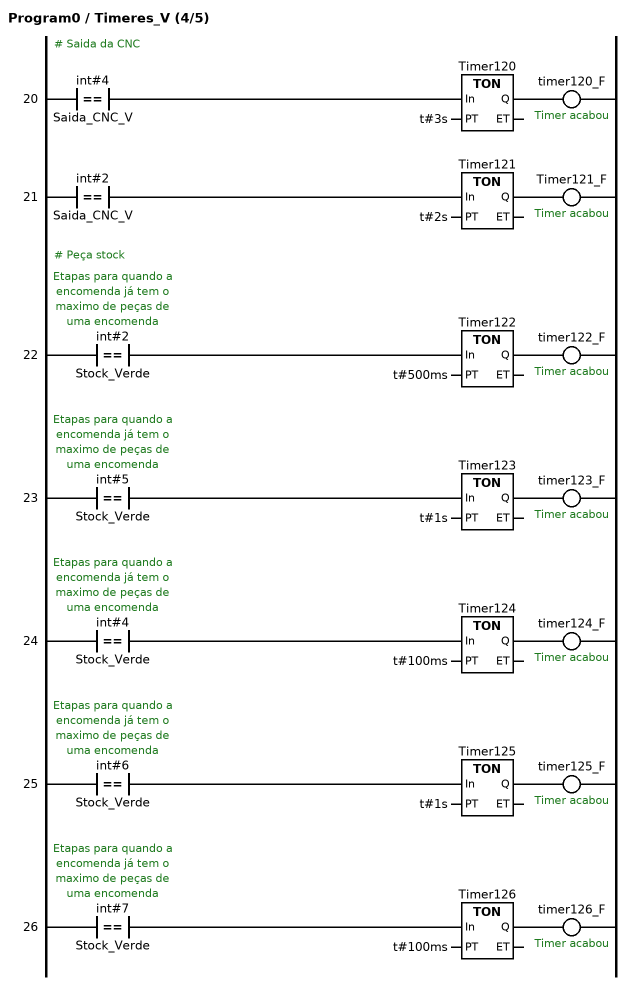
(* [picture p24: Program0 / Timeres_V, rungs 20-26] *)
(* Rung 20: # Saida da CNC *)
Timer120(In := int#4 = Saida_CNC_V, PT := t#3s);
timer120_F := Timer120.Q;
(* Rung 21 *)
Timer121(In := int#2 = Saida_CNC_V, PT := t#2s);
Timer121_F := Timer121.Q;
(* Rung 22: # Peça stock *)
Timer122(In := int#2 = Stock_Verde, PT := t#500ms);
timer122_F := Timer122.Q;
(* Rung 23 *)
Timer123(In := int#5 = Stock_Verde, PT := t#1s);
timer123_F := Timer123.Q;
(* Rung 24 *)
Timer124(In := int#4 = Stock_Verde, PT := t#100ms);
timer124_F := Timer124.Q;
(* Rung 25 *)
Timer125(In := int#6 = Stock_Verde, PT := t#1s);
timer125_F := Timer125.Q;
(* Rung 26 *)
Timer126(In := int#7 = Stock_Verde, PT := t#100ms);
timer126_F := Timer126.Q;

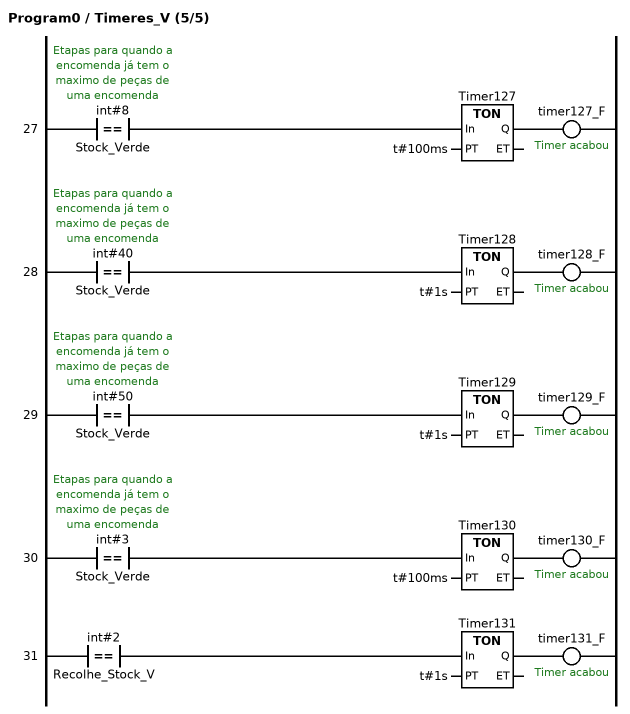
(* Rung 27 *)
Timer127(In := int#8 = Stock_Verde, PT := t#100ms);
timer127_F := Timer127.Q;
(* Rung 28 *)
Timer128(In := int#40 = Stock_Verde, PT := t#1s);
timer128_F := Timer128.Q;
(* Rung 29 *)
Timer129(In := int#50 = Stock_Verde, PT := t#1s);
timer129_F := Timer129.Q;
(* Rung 30 *)
Timer130(In := int#3 = Stock_Verde, PT := t#100ms);
timer130_F := Timer130.Q;
(* Rung 31 *)
Timer131(In := int#2 = Recolhe_Stock_V, PT := t#1s);
timer131_F := Timer131.Q;

(* Section Timeres_C: ladder, written here as Structured Text *)

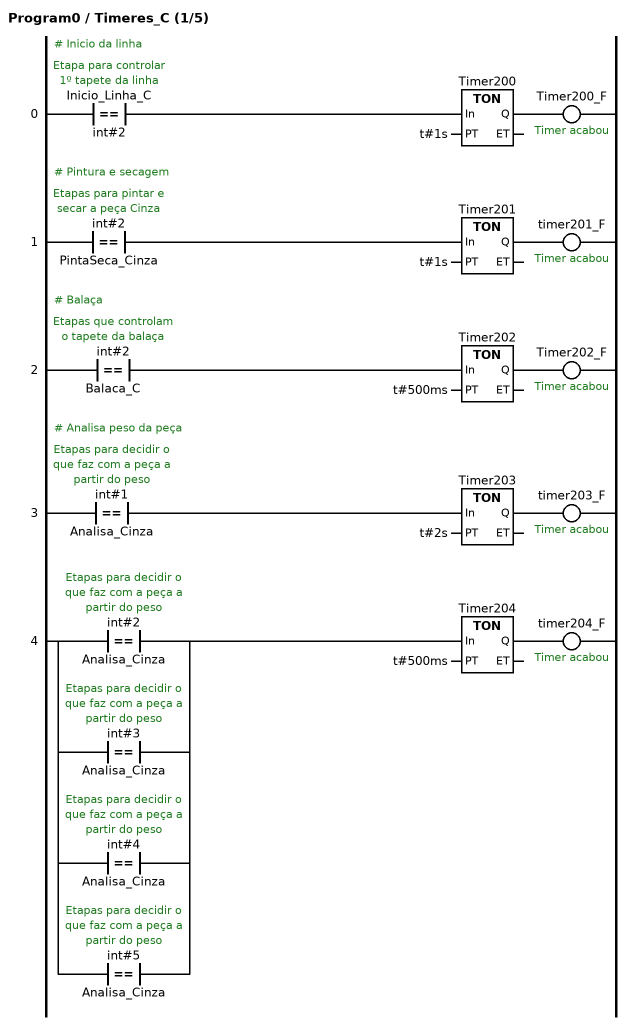
(* Rung 0: # Inicio da linha *)
Timer200(In := Inicio_Linha_C = int#2, PT := t#1s);
Timer200_F := Timer200.Q;
(* Rung 1: # Pintura e secagem *)
Timer201(In := int#2 = PintaSeca_Cinza, PT := t#1s);
timer201_F := Timer201.Q;
(* Rung 2: # Balaça *)
Timer202(In := int#2 = Balaca_C, PT := t#500ms);
Timer202_F := Timer202.Q;
(* Rung 3: # Analisa peso da peça *)
Timer203(In := int#1 = Analisa_Cinza, PT := t#2s);
timer203_F := Timer203.Q;
(* Rung 4 *)
Timer204(In := (int#2 = Analisa_Cinza) OR (int#3 = Analisa_Cinza) OR (int#4 = Analisa_Cinza) OR (int#5 = Analisa_Cinza), PT := t#500ms);
timer204_F := Timer204.Q;

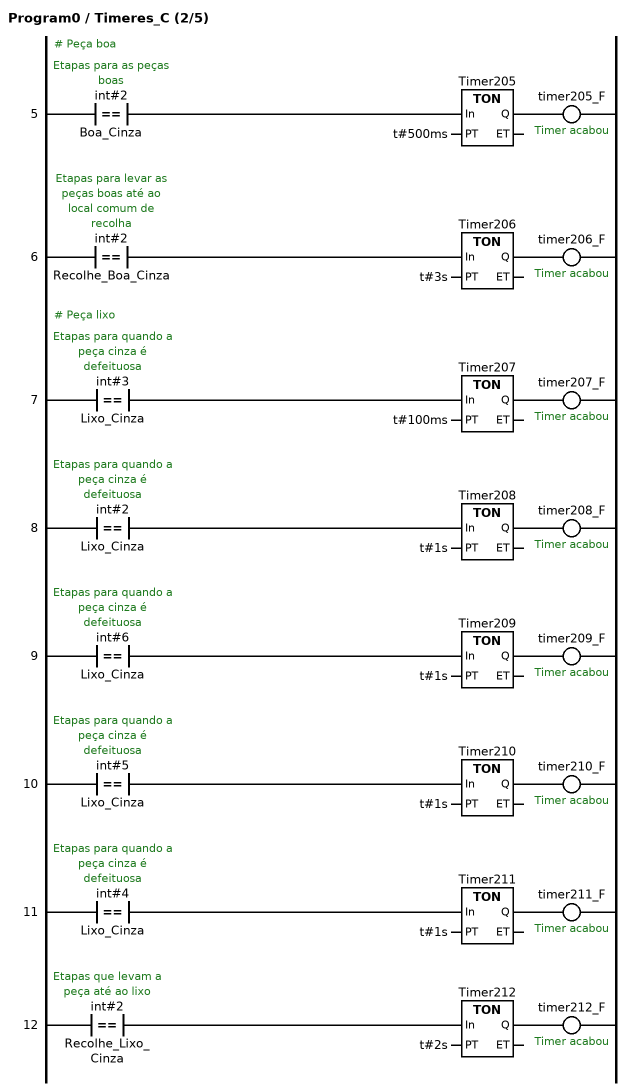
(* Rung 5: # Peça boa *)
Timer205(In := int#2 = Boa_Cinza, PT := t#500ms);
timer205_F := Timer205.Q;
(* Rung 6 *)
Timer206(In := int#2 = Recolhe_Boa_Cinza, PT := t#3s);
timer206_F := Timer206.Q;
(* Rung 7: # Peça lixo *)
Timer207(In := int#3 = Lixo_Cinza, PT := t#100ms);
timer207_F := Timer207.Q;
(* Rung 8 *)
Timer208(In := int#2 = Lixo_Cinza, PT := t#1s);
timer208_F := Timer208.Q;
(* Rung 9 *)
Timer209(In := int#6 = Lixo_Cinza, PT := t#1s);
timer209_F := Timer209.Q;
(* Rung 10 *)
Timer210(In := int#5 = Lixo_Cinza, PT := t#1s);
timer210_F := Timer210.Q;
(* Rung 11 *)
Timer211(In := int#4 = Lixo_Cinza, PT := t#1s);
timer211_F := Timer211.Q;
(* Rung 12 *)
Timer212(In := int#2 = Recolhe_Lixo_Cinza, PT := t#2s);
timer212_F := Timer212.Q;

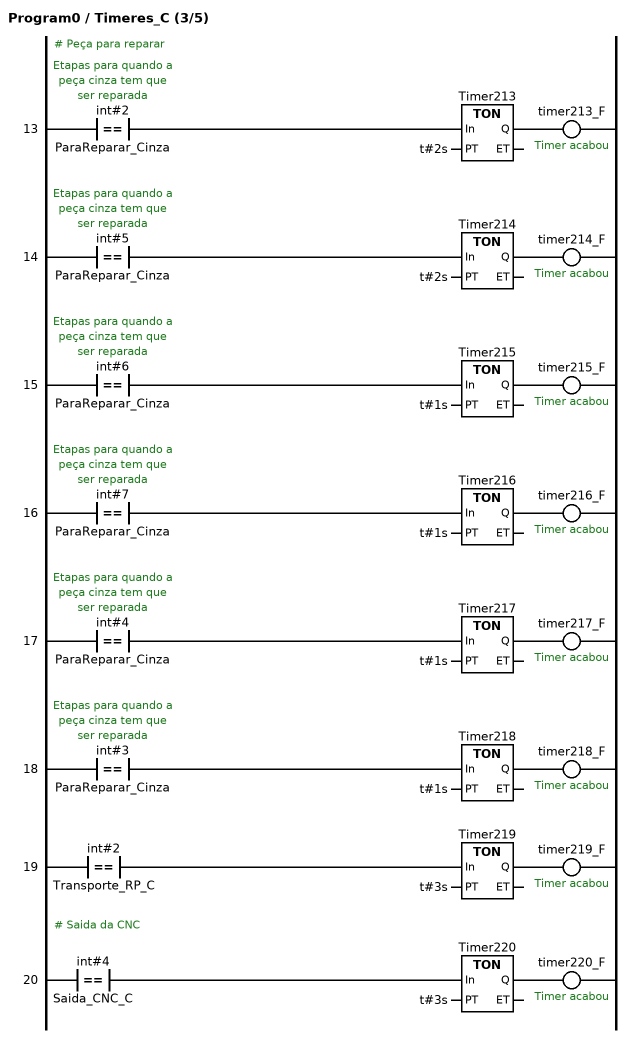
(* Rung 13: # Peça para reparar *)
Timer213(In := int#2 = ParaReparar_Cinza, PT := t#2s);
timer213_F := Timer213.Q;
(* Rung 14 *)
Timer214(In := int#5 = ParaReparar_Cinza, PT := t#2s);
timer214_F := Timer214.Q;
(* Rung 15 *)
Timer215(In := int#6 = ParaReparar_Cinza, PT := t#1s);
timer215_F := Timer215.Q;
(* Rung 16 *)
Timer216(In := int#7 = ParaReparar_Cinza, PT := t#1s);
timer216_F := Timer216.Q;
(* Rung 17 *)
Timer217(In := int#4 = ParaReparar_Cinza, PT := t#1s);
timer217_F := Timer217.Q;
(* Rung 18 *)
Timer218(In := int#3 = ParaReparar_Cinza, PT := t#1s);
timer218_F := Timer218.Q;
(* Rung 19 *)
Timer219(In := int#2 = Transporte_RP_C, PT := t#3s);
timer219_F := Timer219.Q;
(* Rung 20: # Saida da CNC *)
Timer220(In := int#4 = Saida_CNC_C, PT := t#3s);
timer220_F := Timer220.Q;

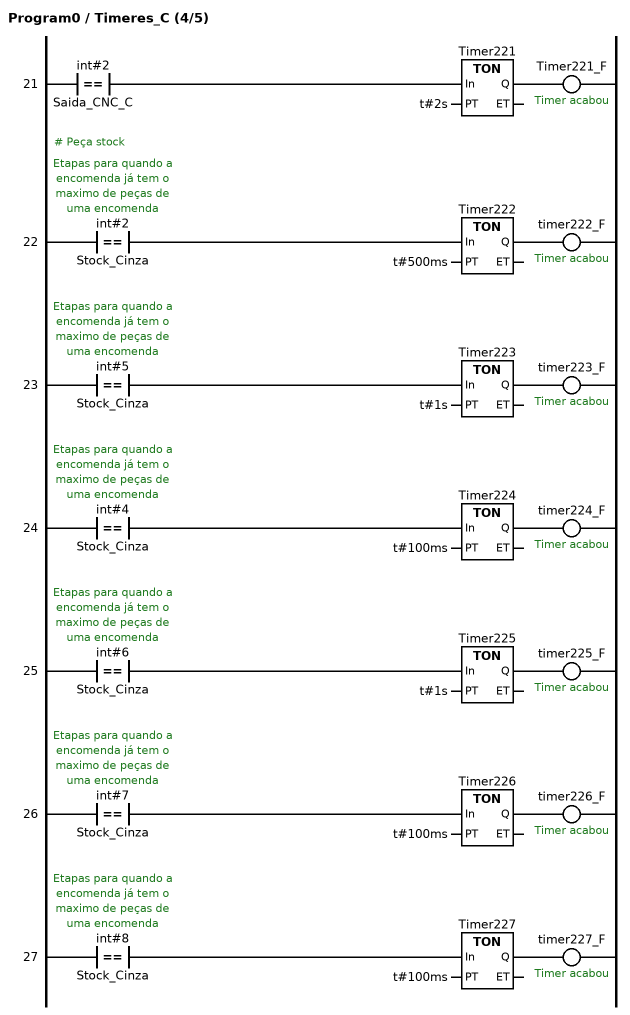
(* Rung 21 *)
Timer221(In := int#2 = Saida_CNC_C, PT := t#2s);
Timer221_F := Timer221.Q;
(* Rung 22: # Peça stock *)
Timer222(In := int#2 = Stock_Cinza, PT := t#500ms);
timer222_F := Timer222.Q;
(* Rung 23 *)
Timer223(In := int#5 = Stock_Cinza, PT := t#1s);
timer223_F := Timer223.Q;
(* Rung 24 *)
Timer224(In := int#4 = Stock_Cinza, PT := t#100ms);
timer224_F := Timer224.Q;
(* Rung 25 *)
Timer225(In := int#6 = Stock_Cinza, PT := t#1s);
timer225_F := Timer225.Q;
(* Rung 26 *)
Timer226(In := int#7 = Stock_Cinza, PT := t#100ms);
timer226_F := Timer226.Q;
(* Rung 27 *)
Timer227(In := int#8 = Stock_Cinza, PT := t#100ms);
timer227_F := Timer227.Q;

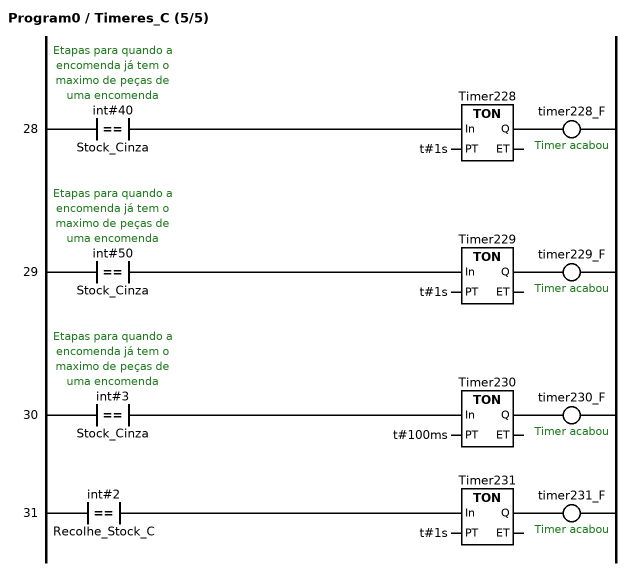
(* Rung 28 *)
Timer228(In := int#40 = Stock_Cinza, PT := t#1s);
timer228_F := Timer228.Q;
(* Rung 29 *)
Timer229(In := int#50 = Stock_Cinza, PT := t#1s);
timer229_F := Timer229.Q;
(* Rung 30 *)
Timer230(In := int#3 = Stock_Cinza, PT := t#100ms);
timer230_F := Timer230.Q;
(* Rung 31 *)
Timer231(In := int#2 = Recolhe_Stock_C, PT := t#1s);
timer231_F := Timer231.Q;

(* Section Emitter_Removers: ladder, written here as Structured Text *)

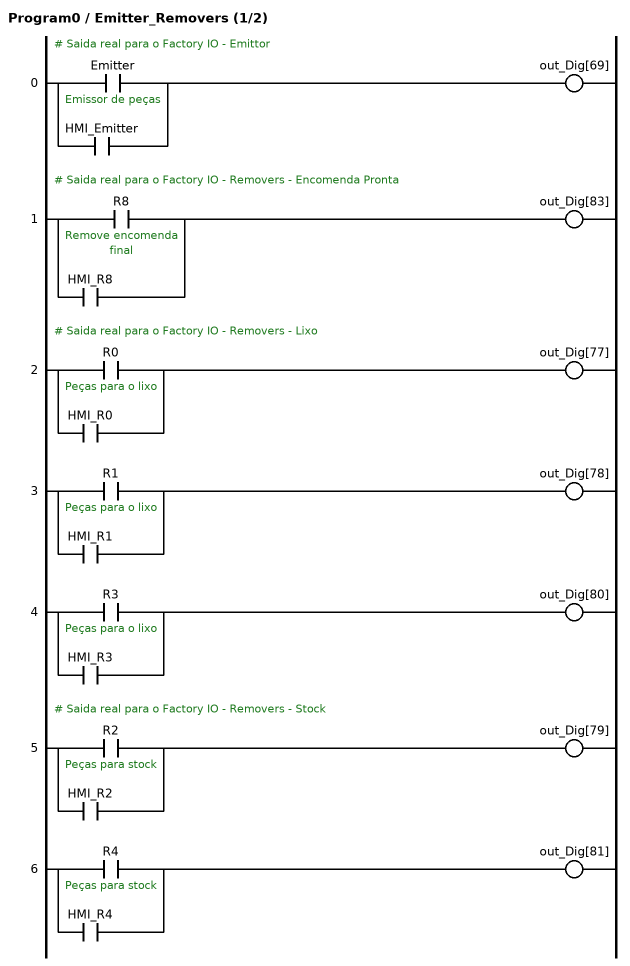
(* Rung 0: # Saida real para o Factory IO - Emittor *)
out_Dig[69] := Emitter OR HMI_Emitter;
(* Rung 1: # Saida real para o Factory IO - Removers - Encomenda Pronta *)
out_Dig[83] := R8 OR HMI_R8;
(* Rung 2: # Saida real para o Factory IO - Removers - Lixo *)
out_Dig[77] := R0 OR HMI_R0;
(* Rung 3 *)
out_Dig[78] := R1 OR HMI_R1;
(* Rung 4 *)
out_Dig[80] := R3 OR HMI_R3;
(* Rung 5: # Saida real para o Factory IO - Removers - Stock *)
out_Dig[79] := R2 OR HMI_R2;
(* Rung 6 *)
out_Dig[81] := R4 OR HMI_R4;

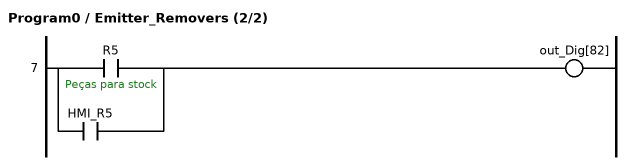
(* Rung 7 *)
out_Dig[82] := R5 OR HMI_R5;

(* Section Semaforos_Alarme: ladder, written here as Structured Text *)

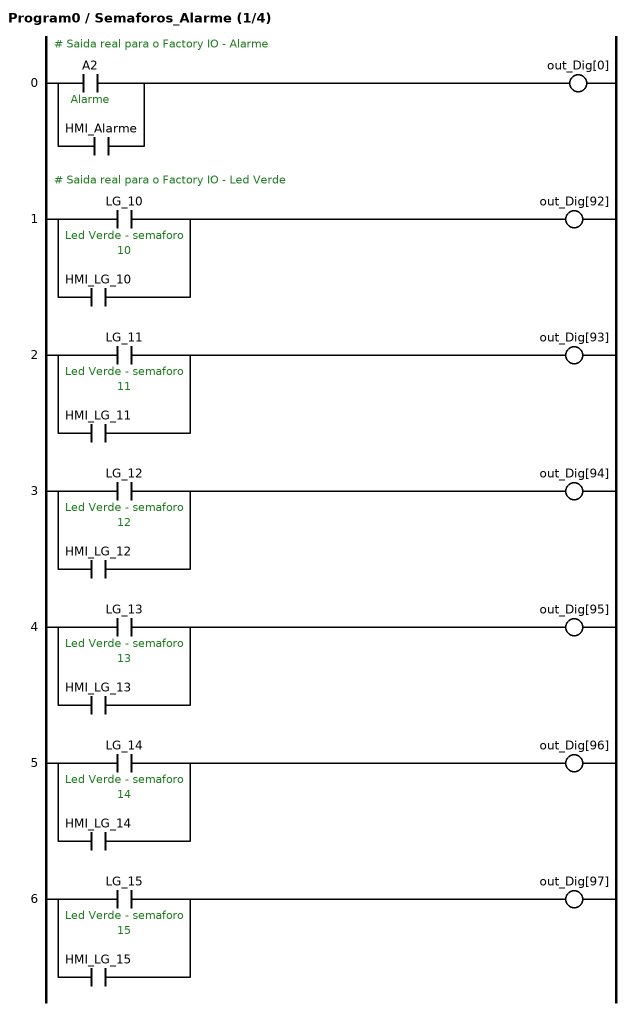
(* Rung 0: # Saida real para o Factory IO - Alarme *)
out_Dig[0] := A2 OR HMI_Alarme;
(* Rung 1: # Saida real para o Factory IO - Led Verde *)
out_Dig[92] := LG_10 OR HMI_LG_10;
(* Rung 2 *)
out_Dig[93] := LG_11 OR HMI_LG_11;
(* Rung 3 *)
out_Dig[94] := LG_12 OR HMI_LG_12;
(* Rung 4 *)
out_Dig[95] := LG_13 OR HMI_LG_13;
(* Rung 5 *)
out_Dig[96] := LG_14 OR HMI_LG_14;
(* Rung 6 *)
out_Dig[97] := LG_15 OR HMI_LG_15;

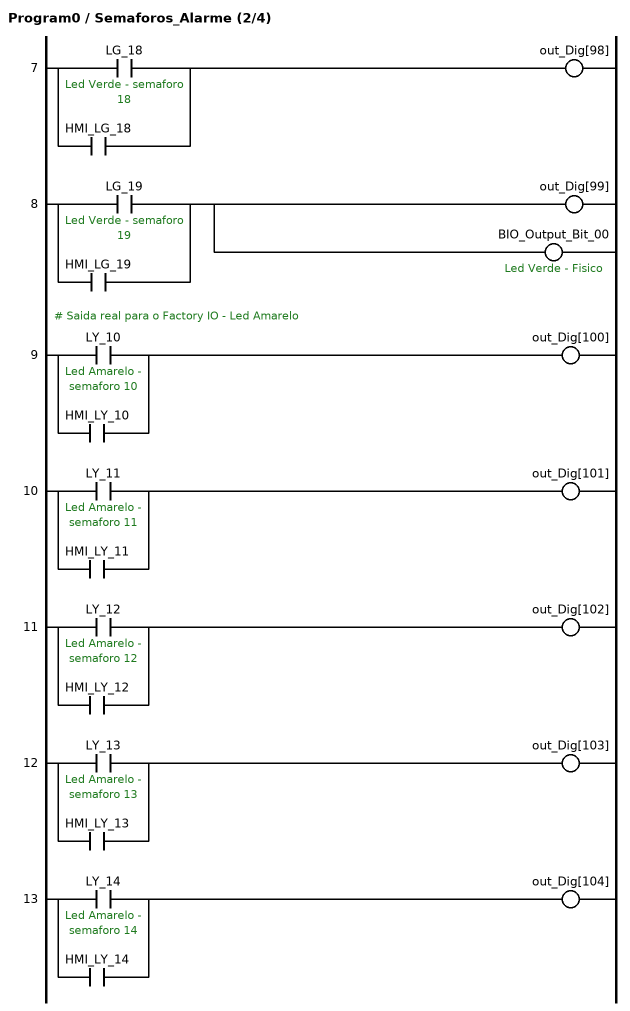
(* Rung 7 *)
out_Dig[98] := LG_18 OR HMI_LG_18;
(* Rung 8 *)
out_Dig[99] := LG_19 OR HMI_LG_19;
BIO_Output_Bit_00 := LG_19 OR HMI_LG_19;
(* Rung 9: # Saida real para o Factory IO - Led Amarelo *)
out_Dig[100] := LY_10 OR HMI_LY_10;
(* Rung 10 *)
out_Dig[101] := LY_11 OR HMI_LY_11;
(* Rung 11 *)
out_Dig[102] := LY_12 OR HMI_LY_12;
(* Rung 12 *)
out_Dig[103] := LY_13 OR HMI_LY_13;
(* Rung 13 *)
out_Dig[104] := LY_14 OR HMI_LY_14;

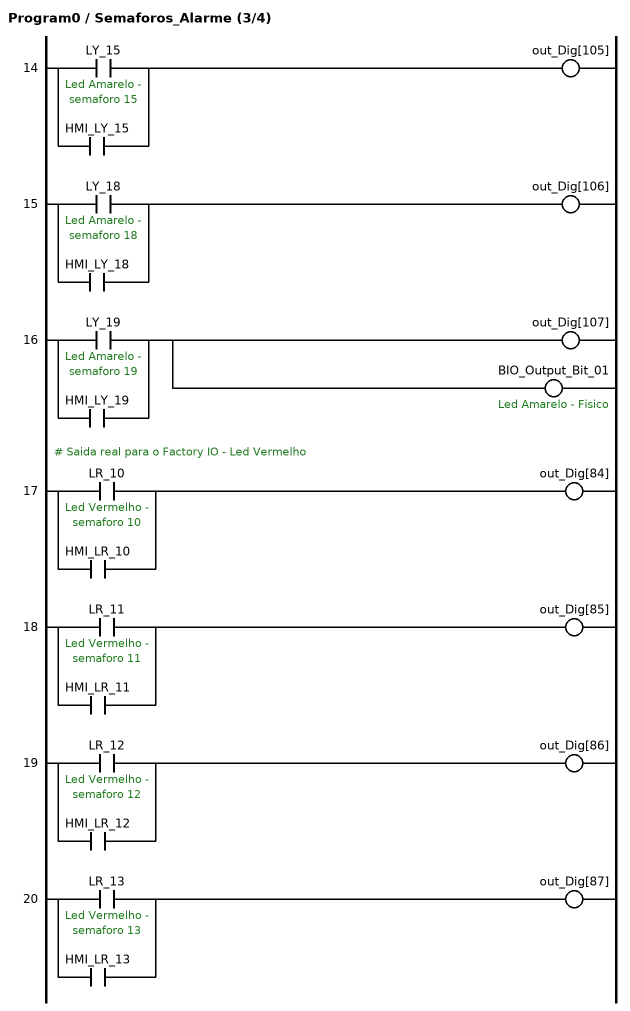
(* Rung 14 *)
out_Dig[105] := LY_15 OR HMI_LY_15;
(* Rung 15 *)
out_Dig[106] := LY_18 OR HMI_LY_18;
(* Rung 16 *)
out_Dig[107] := LY_19 OR HMI_LY_19;
BIO_Output_Bit_01 := LY_19 OR HMI_LY_19;
(* Rung 17: # Saida real para o Factory IO - Led Vermelho *)
out_Dig[84] := LR_10 OR HMI_LR_10;
(* Rung 18 *)
out_Dig[85] := LR_11 OR HMI_LR_11;
(* Rung 19 *)
out_Dig[86] := LR_12 OR HMI_LR_12;
(* Rung 20 *)
out_Dig[87] := LR_13 OR HMI_LR_13;

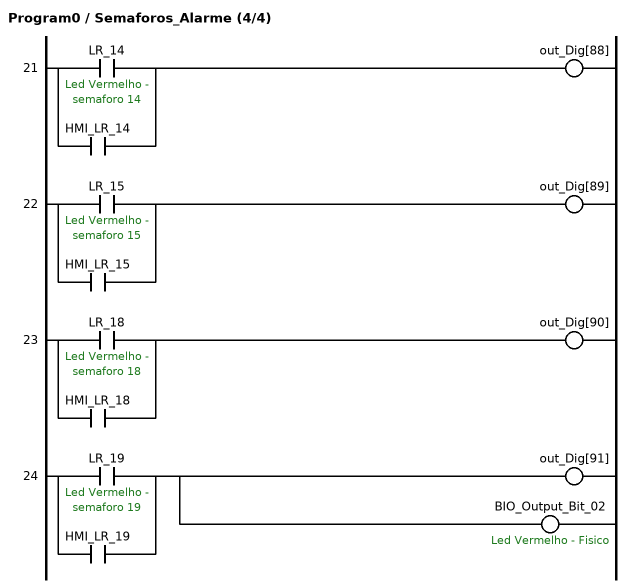
(* Rung 21 *)
out_Dig[88] := LR_14 OR HMI_LR_14;
(* Rung 22 *)
out_Dig[89] := LR_15 OR HMI_LR_15;
(* Rung 23 *)
out_Dig[90] := LR_18 OR HMI_LR_18;
(* Rung 24 *)
out_Dig[91] := LR_19 OR HMI_LR_19;
BIO_Output_Bit_02 := LR_19 OR HMI_LR_19;

(* Section Pick_and_Place: ladder, written here as Structured Text *)

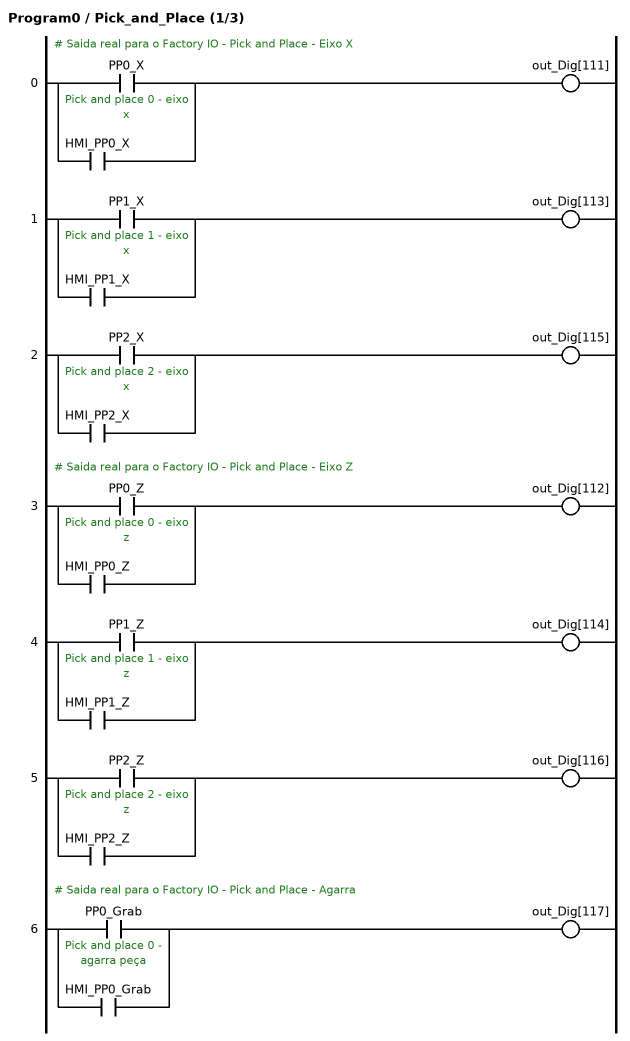
(* Rung 0: # Saida real para o Factory IO - Pick and Place - Eixo X *)
out_Dig[111] := PP0_X OR HMI_PP0_X;
(* Rung 1 *)
out_Dig[113] := PP1_X OR HMI_PP1_X;
(* Rung 2 *)
out_Dig[115] := PP2_X OR HMI_PP2_X;
(* Rung 3: # Saida real para o Factory IO - Pick and Place - Eixo Z *)
out_Dig[112] := PP0_Z OR HMI_PP0_Z;
(* Rung 4 *)
out_Dig[114] := PP1_Z OR HMI_PP1_Z;
(* Rung 5 *)
out_Dig[116] := PP2_Z OR HMI_PP2_Z;
(* Rung 6: # Saida real para o Factory IO - Pick and Place - Agarra *)
out_Dig[117] := PP0_Grab OR HMI_PP0_Grab;

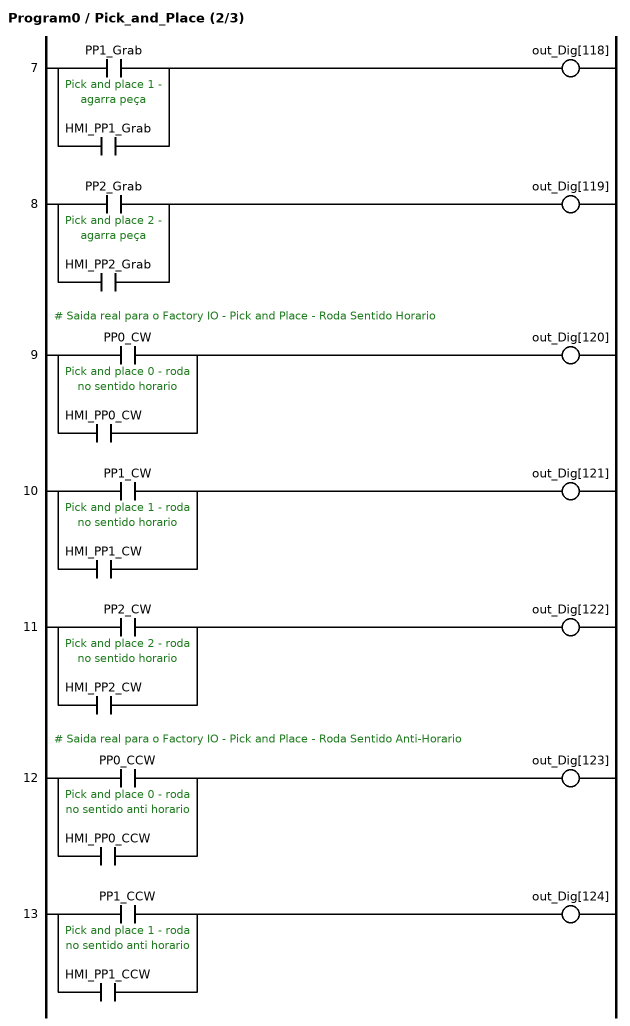
(* Rung 7 *)
out_Dig[118] := PP1_Grab OR HMI_PP1_Grab;
(* Rung 8 *)
out_Dig[119] := PP2_Grab OR HMI_PP2_Grab;
(* Rung 9: # Saida real para o Factory IO - Pick and Place - Roda Sentido Horario *)
out_Dig[120] := PP0_CW OR HMI_PP0_CW;
(* Rung 10 *)
out_Dig[121] := PP1_CW OR HMI_PP1_CW;
(* Rung 11 *)
out_Dig[122] := PP2_CW OR HMI_PP2_CW;
(* Rung 12: # Saida real para o Factory IO - Pick and Place - Roda Sentido Anti-Horario *)
out_Dig[123] := PP0_CCW OR HMI_PP0_CCW;
(* Rung 13 *)
out_Dig[124] := PP1_CCW OR HMI_PP1_CCW;

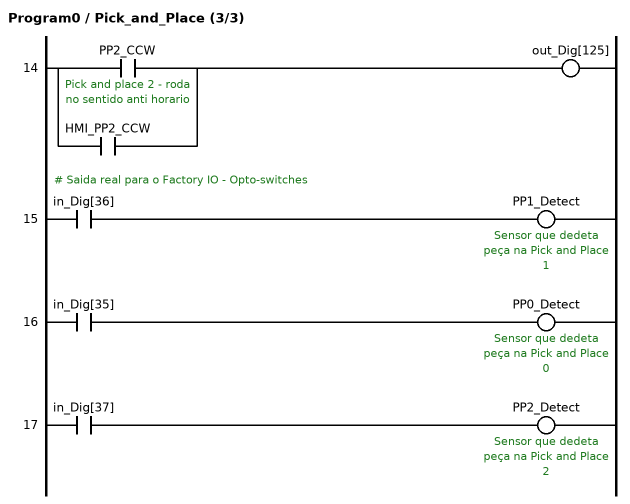
(* Rung 14 *)
out_Dig[125] := PP2_CCW OR HMI_PP2_CCW;
(* Rung 15: # Saida real para o Factory IO - Opto-switches *)
PP1_Detect := in_Dig[36];
(* Rung 16 *)
PP0_Detect := in_Dig[35];
(* Rung 17 *)
PP2_Detect := in_Dig[37];

(* Section Pick_and_Place_0_S: ladder, written here as Structured Text *)

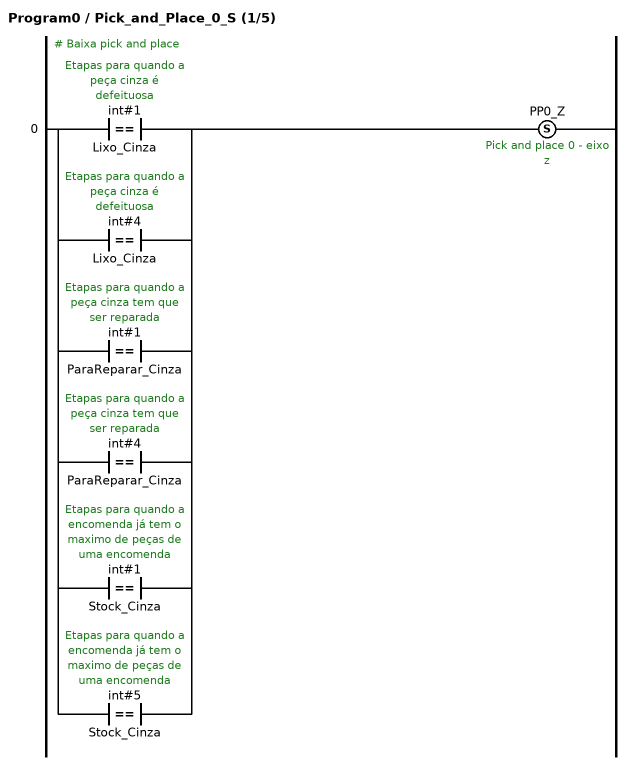
(* Rung 0: # Baixa pick and place *)
IF (int#1 = Lixo_Cinza) OR (int#4 = Lixo_Cinza) OR (int#1 = ParaReparar_Cinza) OR (int#4 = ParaReparar_Cinza) OR (int#1 = Stock_Cinza) OR (int#5 = Stock_Cinza) THEN
    PP0_Z := TRUE;
END_IF;

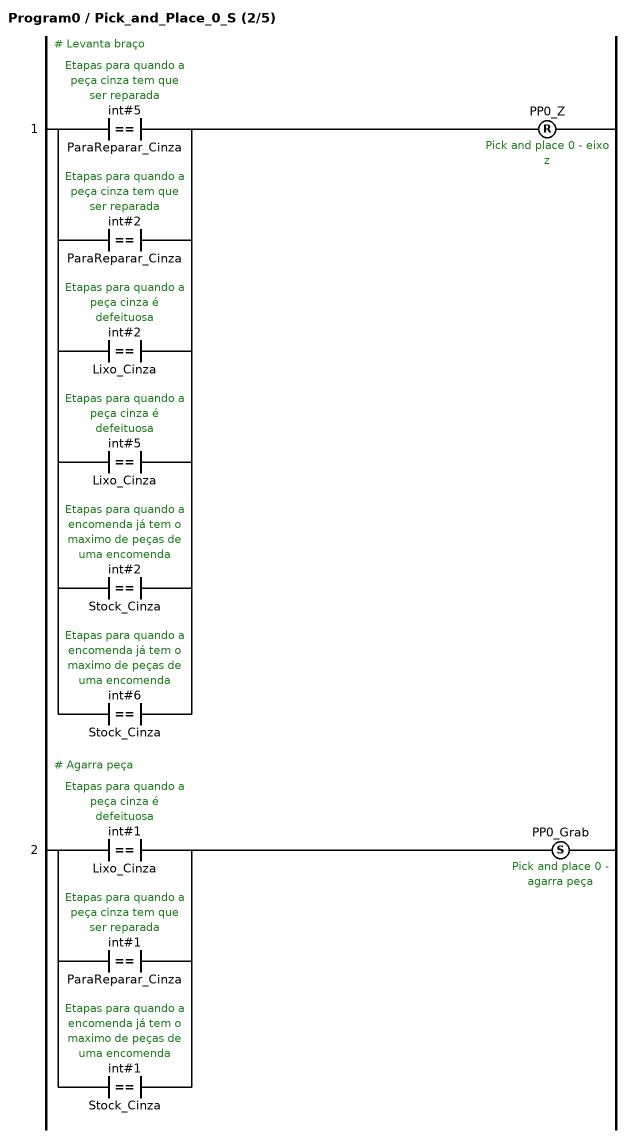
(* Rung 1: # Levanta braço *)
IF (int#5 = ParaReparar_Cinza) OR (int#2 = ParaReparar_Cinza) OR (int#2 = Lixo_Cinza) OR (int#5 = Lixo_Cinza) OR (int#2 = Stock_Cinza) OR (int#6 = Stock_Cinza) THEN
    PP0_Z := FALSE;
END_IF;
(* Rung 2: # Agarra peça *)
IF (int#1 = Lixo_Cinza) OR (int#1 = ParaReparar_Cinza) OR (int#1 = Stock_Cinza) THEN
    PP0_Grab := TRUE;
END_IF;

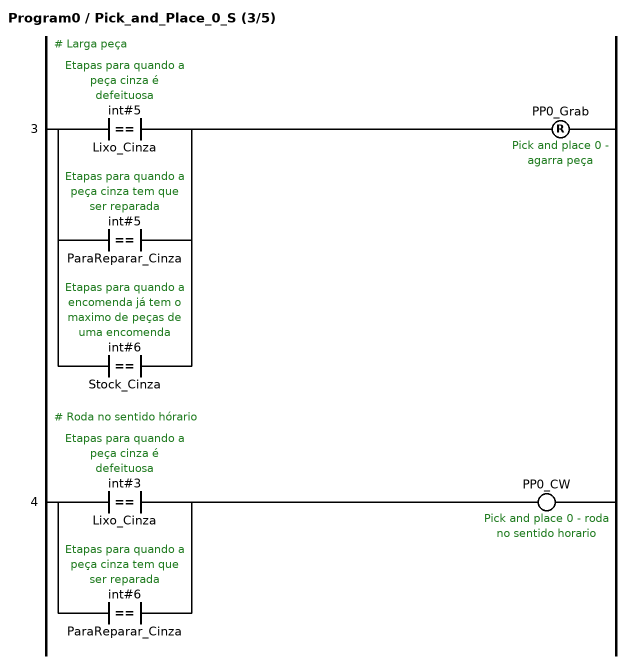
(* Rung 3: # Larga peça *)
IF (int#5 = Lixo_Cinza) OR (int#5 = ParaReparar_Cinza) OR (int#6 = Stock_Cinza) THEN
    PP0_Grab := FALSE;
END_IF;
(* Rung 4: # Roda no sentido hórario *)
PP0_CW := (int#3 = Lixo_Cinza) OR (int#6 = ParaReparar_Cinza);

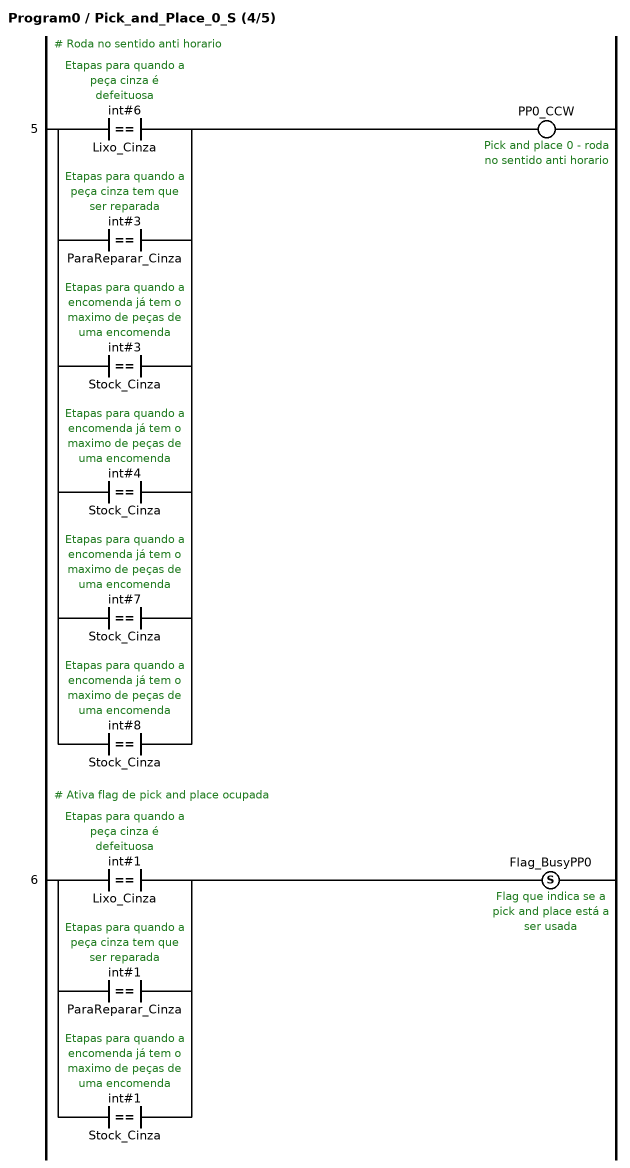
(* Rung 5: # Roda no sentido anti horario *)
PP0_CCW := (int#6 = Lixo_Cinza) OR (int#3 = ParaReparar_Cinza) OR (int#3 = Stock_Cinza) OR (int#4 = Stock_Cinza) OR (int#7 = Stock_Cinza) OR (int#8 = Stock_Cinza);
(* Rung 6: # Ativa flag de pick and place ocupada *)
IF (int#1 = Lixo_Cinza) OR (int#1 = ParaReparar_Cinza) OR (int#1 = Stock_Cinza) THEN
    Flag_BusyPP0 := TRUE;
END_IF;

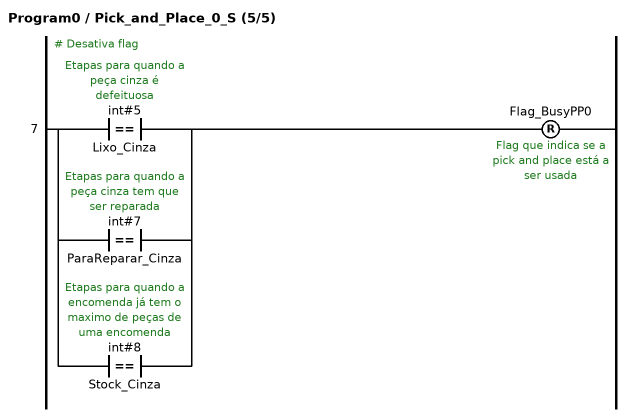
(* Rung 7: # Desativa flag *)
IF (int#5 = Lixo_Cinza) OR (int#7 = ParaReparar_Cinza) OR (int#8 = Stock_Cinza) THEN
    Flag_BusyPP0 := FALSE;
END_IF;

(* Section Pick_and_Place_1_S: ladder, written here as Structured Text *)

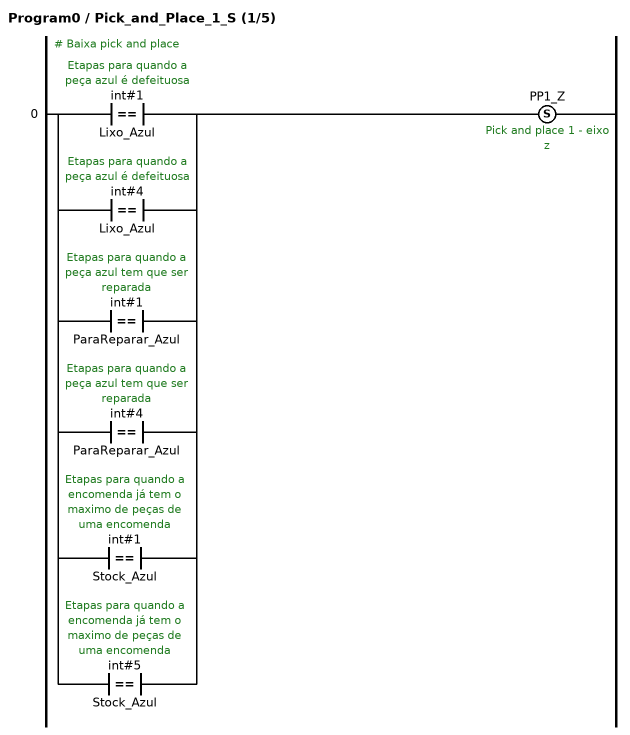
(* Rung 0: # Baixa pick and place *)
IF (int#1 = Lixo_Azul) OR (int#4 = Lixo_Azul) OR (int#1 = ParaReparar_Azul) OR (int#4 = ParaReparar_Azul) OR (int#1 = Stock_Azul) OR (int#5 = Stock_Azul) THEN
    PP1_Z := TRUE;
END_IF;

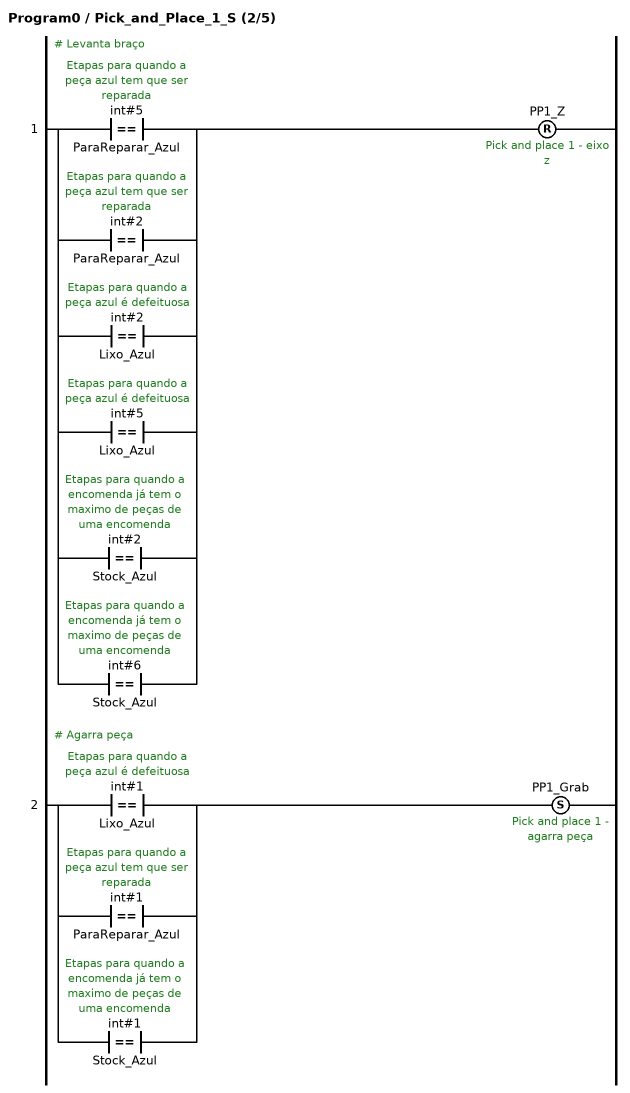
(* Rung 1: # Levanta braço *)
IF (int#5 = ParaReparar_Azul) OR (int#2 = ParaReparar_Azul) OR (int#2 = Lixo_Azul) OR (int#5 = Lixo_Azul) OR (int#2 = Stock_Azul) OR (int#6 = Stock_Azul) THEN
    PP1_Z := FALSE;
END_IF;
(* Rung 2: # Agarra peça *)
IF (int#1 = Lixo_Azul) OR (int#1 = ParaReparar_Azul) OR (int#1 = Stock_Azul) THEN
    PP1_Grab := TRUE;
END_IF;

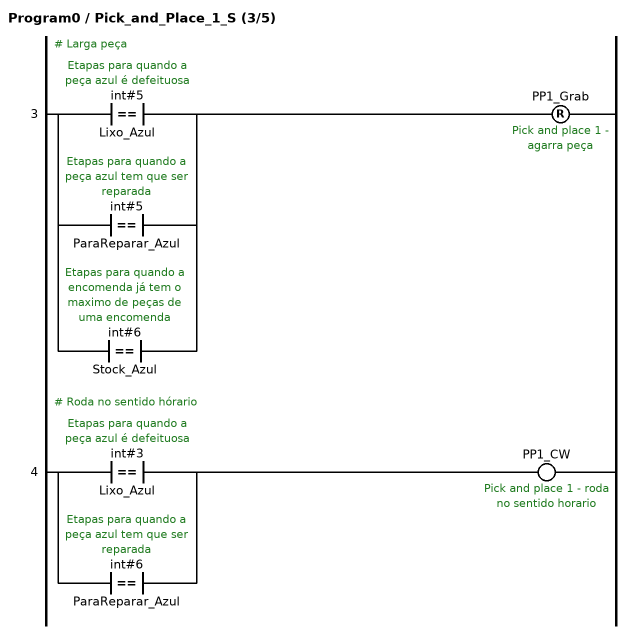
(* Rung 3: # Larga peça *)
IF (int#5 = Lixo_Azul) OR (int#5 = ParaReparar_Azul) OR (int#6 = Stock_Azul) THEN
    PP1_Grab := FALSE;
END_IF;
(* Rung 4: # Roda no sentido hórario *)
PP1_CW := (int#3 = Lixo_Azul) OR (int#6 = ParaReparar_Azul);

